FUNCTION_BLOCK DRIVE
  VAR_INPUT
    Start : BOOL;
    Stop  : BOOL;
  END_VAR
  VAR_OUTPUT
    Run : BOOL;
  END_VAR

BEGIN
Run := (Start OR Run) AND NOT Stop;
  //#ASSERT NOT Run OR NOT Stop : P1
END_FUNCTION_BLOCK
